(* IEC 61131-3 sources: SemaPLC/sema-plc-benchmark/spec2control-benchmark/data/st-baseline/coking-refinery/pous/programs, 9 files *)

(* ---- main.st ---- *)
PROGRAM main
VAR
	Heartbeat : bool;
END_VAR

(* Entry point required by OpenPLC Editor v4. The process sections run as parallel program instances under task0; main only provides a scan heartbeat. *)
Heartbeat := NOT Heartbeat;

END_PROGRAM

(* ---- Section2.st ---- *)
PROGRAM Section2
VAR
	FT101_FeedFlow_PV_kgphr : real;
	FT102_RefluxFlow_PV_kgphr : real;
	FFIC103_RefluxFlow_SP_kgphr : real;
	FIC104_Output_Percent : real;
	FV104_ValvePosition_Percent : real;
	FV104_FeedbackPos_Percent : real;
	FV104_ValveMoving : bool;
	PIT106_ColumnPressure_bar : real;
	TIT104_Temperature_C : real;
	TIT105_Temperature_C : real;
	TIT107_Temperature_C : real;
	FT_101 : ANALOG_IN;
	FT_102 : ANALOG_IN;
	PIT_106 : ANALOG_IN;
	TIT_104 : ANALOG_IN;
	TIT_105 : ANALOG_IN;
	TIT_107 : ANALOG_IN;
	FFIC_103 : RATIO_CONTROL;
	FIC_104 : PID_BASIC;
	FV_104 : VALVE_ELECTRIC;
	RatioInhibit_OR : bool;
	FeedNotAbove500_NOT : bool;
	ValveInhibit_OR : bool;
END_VAR

FT_101(
    PV_Low := 100.0,
    Scaling_Slope := 312.5,
    Scaling_Offset := -1250.0,
    Alarm_Enable := TRUE);
FT_102(
    Scaling_Slope := 156.25,
    Scaling_Offset := -625.0,
    Alarm_Enable := TRUE);
PIT_106(
    PV_High := 1.5,
    PV_Low := 0.5,
    Alarm_Enable := TRUE);
TIT_104(
    PV_High := 350.0,
    PV_Low := 120.0,
    Alarm_Enable := TRUE);
TIT_105(
    PV_High := 350.0,
    PV_Low := 120.0,
    Alarm_Enable := TRUE);
TIT_107(
    PV_High := 350.0,
    PV_Low := 120.0,
    Alarm_Enable := TRUE);
FIC_104(
    AUTO := TRUE,
    PV := FT_102.PV,
    SP := FFIC_103.SlaveSP,
    MV_MIN := 0.0,
    MV_MAX := 100.0,
    Inhibit := RatioInhibit_OR);
FeedNotAbove500_NOT := NOT FT_101.High_Alarm;
ValveInhibit_OR := FeedNotAbove500_NOT OR TIT_104.High_Alarm OR TIT_104.Low_Alarm OR TIT_105.High_Alarm OR TIT_105.Low_Alarm OR TIT_107.High_Alarm OR TIT_107.Low_Alarm;
FV_104(
    Control_Signal := FIC_104.XOUT,
    Manual_Mode := FALSE,
    Open_Limit := 100.0,
    Close_Limit := 0.0,
    Inhibit := ValveInhibit_OR);
RatioInhibit_OR := PIT_106.High_Alarm OR PIT_106.Low_Alarm OR TIT_104.High_Alarm OR TIT_104.Low_Alarm OR TIT_105.High_Alarm OR TIT_105.Low_Alarm OR TIT_107.High_Alarm OR TIT_107.Low_Alarm OR FT_101.Low_Alarm OR FT_101.General_Fault OR FT_102.General_Fault OR FV_104.Position_Error;
FFIC_103(
    Auto := TRUE,
    PrimaryPV := FT_101.PV,
    SecondaryPV := FT_102.PV,
    RatioSP := 0.5,
    Bias := 0.0,
    MV_MIN := 0.0,
    MV_MAX := 2500.0,
    Inhibit := RatioInhibit_OR);

(* Outputs published to other sections / HMI. *)
FT101_FeedFlow_PV_kgphr := FT_101.PV;
FT102_RefluxFlow_PV_kgphr := FT_102.PV;
FFIC103_RefluxFlow_SP_kgphr := FFIC_103.SlaveSP;
FIC104_Output_Percent := FIC_104.XOUT;
FV104_ValvePosition_Percent := FV_104.Valve_Position;
FV104_FeedbackPos_Percent := FV_104.Feedback_Pos;
FV104_ValveMoving := FV_104.Valve_Moving;
PIT106_ColumnPressure_bar := PIT_106.PV;
TIT104_Temperature_C := TIT_104.PV;
TIT105_Temperature_C := TIT_105.PV;
TIT107_Temperature_C := TIT_107.PV;

END_PROGRAM

(* ---- Section3.st ---- *)
PROGRAM Section3
VAR
	PIT_103_PV_mmHg : real;
	PIC_102_MV_Percent : real;
	PIT_103 : ANALOG_IN;
	PIC_102 : PID_BASIC;
	PV_101 : VALVE_ELECTRIC;
	VDU_START_OK : BOOL_INPUT;
	MAINT_BYPASS_OK : BOOL_INPUT;
	PIC102Inhibit_OR : bool;
	PV101Inhibit_OR : bool;
	VDUStartPermissive_NOT : bool;
END_VAR

PIT_103(
    PV_High := 80.0,
    PV_Low := 20.0,
    Scaling_Slope := 47.5,
    Scaling_Offset := -190.0,
    Alarm_Enable := TRUE);
MAINT_BYPASS_OK();
VDU_START_OK();
VDUStartPermissive_NOT := NOT VDU_START_OK.Bool_Out;
PIC102Inhibit_OR := VDUStartPermissive_NOT OR MAINT_BYPASS_OK.Bool_Out OR PIT_103.General_Fault OR PIC_102.PV_Low_Alarm;
PIC_102(
    AUTO := TRUE,
    PV := PIT_103.PV,
    SP := 50.0,
    MV_MIN := 0.0,
    MV_MAX := 100.0,
    KP := 1.8,
    TR := 2.0,
    TD := 0.5,
    Deviation_Limit := 5.0,
    Inhibit := PIC102Inhibit_OR);
PV101Inhibit_OR := PIC_102.PV_High_Alarm OR PV_101.Position_Error;
PV_101(
    Control_Signal := PIC_102.XOUT,
    Open_Limit := 100.0,
    Close_Limit := 0.0,
    Inhibit := PV101Inhibit_OR);

(* Outputs published to other sections / HMI. *)
PIT_103_PV_mmHg := PIT_103.PV;
PIC_102_MV_Percent := PIC_102.XOUT;

END_PROGRAM

(* ---- Section4.st ---- *)
PROGRAM Section4
VAR
	PC301_SP_Operator : real;
	PT_301_RegeneratorPressure_PV : real;
	PT_302_BlowerDischargePressure_PV : real;
	PT_303_FractionatorOverheadPressure_PV : real;
	TT_301_RegeneratorTemperature_PV : real;
	PTF_301_FilteredPressure_PV : real;
	PC_301_Output_to_PV_105_Percent : real;
	PV_105_Valve_Position_Command_Percent : real;
	PV_105_Valve_Position_Feedback_Percent : real;
	P_301A_Running_Status : bool;
	XV_108_Closed_Status : bool;
	PT_301 : ANALOG_IN;
	PT_302 : ANALOG_IN;
	PT_303 : ANALOG_IN;
	PTF_301 : ANALOG_IN;
	TT_301 : ANALOG_IN;
	PC_301 : PID_BASIC;
	PV_105 : VALVE_ELECTRIC;
	PV_106 : VALVE_ON_OFF;
	XV_108 : VALVE_ON_OFF;
	P_301A : MOTOR_ON_OFF;
	SteadyState_TON : TON;
	SetpointClamp_LIMIT : real;
	StartupSP_Select_SEL : real;
	ErrorCalc_SUB : real;
	ErrorPos_GT : bool;
	ErrorNeg_LT : bool;
	ErrorOutsideBand_OR : bool;
	DeadbandApply_SEL : real;
	PV_Reconstruct_ADD : real;
	BlowerNotRunning_NOT : bool;
	Permissives_OR1 : bool;
	Permissives_OR2 : bool;
	Permissives_OR3 : bool;
	PV105Inhibit_OR : bool;
	AutoHold_OR : bool;
	AutoEnable_NOT : bool;
	ESD_HighPressure_GT : bool;
	ReliefValve_GT : bool;
	ReliefValve_Close_NOT : bool;
	OutsideBand_NOT : bool;
END_VAR

PT_301(
    PV_High := 2.8,
    PV_Low := 2.2,
    Scaling_Slope := 0.3125,
    Scaling_Offset := -1.25,
    Alarm_Enable := TRUE);
PT_302(
    Scaling_Slope := 0.3125,
    Scaling_Offset := -1.25,
    Alarm_Enable := TRUE);
PT_303(
    Scaling_Slope := 0.3125,
    Scaling_Offset := -1.25,
    Alarm_Enable := TRUE);
PTF_301(
    Scaling_Slope := 0.3125,
    Scaling_Offset := -1.25);
TT_301(
    Scaling_Slope := 62.5,
    Scaling_Offset := -250.0,
    Alarm_Enable := TRUE);
ESD_HighPressure_GT := (PT_301.PV > 3.0);
XV_108(
    Open_Cmd := FALSE,
    Close_Cmd := ESD_HighPressure_GT,
    Timeout := T#5s);
AutoHold_OR := PT_301.General_Fault OR XV_108.FB_Closed;
AutoEnable_NOT := NOT AutoHold_OR;
ErrorNeg_LT := (ErrorCalc_SUB < -0.05);
ErrorPos_GT := (ErrorCalc_SUB > 0.05);
ErrorOutsideBand_OR := ErrorPos_GT OR ErrorNeg_LT;
OutsideBand_NOT := NOT ErrorOutsideBand_OR;
SteadyState_TON(
    IN := OutsideBand_NOT,
    PT := T#60s);
StartupSP_Select_SEL := SEL(G := SteadyState_TON.Q, IN0 := 2.5, IN1 := 0.0);
ErrorCalc_SUB := PT_301.PV - StartupSP_Select_SEL;
DeadbandApply_SEL := SEL(G := ErrorOutsideBand_OR, IN0 := 0.0, IN1 := ErrorCalc_SUB);
PV_Reconstruct_ADD := StartupSP_Select_SEL + DeadbandApply_SEL;
PC_301(
    AUTO := AutoEnable_NOT,
    PV := PV_Reconstruct_ADD,
    SP := StartupSP_Select_SEL,
    MV_MIN := 0.0,
    MV_MAX := 100.0,
    X0 := 0.0,
    KP := 3.0,
    TR := 1.2,
    TD := 0.1);
P_301A();
BlowerNotRunning_NOT := NOT P_301A.FB_Running;
Permissives_OR1 := TT_301.Low_Alarm OR BlowerNotRunning_NOT;
Permissives_OR2 := PT_302.Low_Alarm OR PT_303.High_Alarm;
Permissives_OR3 := Permissives_OR1 OR Permissives_OR2;
PV105Inhibit_OR := Permissives_OR3 OR XV_108.FB_Closed;
PV_105(
    Control_Signal := PC_301.XOUT,
    Manual_Mode := FALSE,
    Open_Limit := 100.0,
    Close_Limit := 0.0,
    Timeout := T#10s,
    Inhibit := PV105Inhibit_OR);
ReliefValve_GT := (PT_301.PV > 3.5);
ReliefValve_Close_NOT := NOT ReliefValve_GT;
PV_106(
    Open_Cmd := ReliefValve_GT,
    Close_Cmd := ReliefValve_Close_NOT,
    Timeout := T#5s);
SetpointClamp_LIMIT := LIMIT(MN := 2.0, IN := PC301_SP_Operator, MX := 3.0);

(* Outputs published to other sections / HMI. *)
PT_301_RegeneratorPressure_PV := PT_301.PV;
PT_302_BlowerDischargePressure_PV := PT_302.PV;
PT_303_FractionatorOverheadPressure_PV := PT_303.PV;
TT_301_RegeneratorTemperature_PV := TT_301.PV;
PTF_301_FilteredPressure_PV := PTF_301.PV;
PC_301_Output_to_PV_105_Percent := PC_301.XOUT;
PV_105_Valve_Position_Command_Percent := PV_105.Valve_Position;
PV_105_Valve_Position_Feedback_Percent := PV_105.Feedback_Pos;
P_301A_Running_Status := P_301A.FB_Running;
XV_108_Closed_Status := XV_108.FB_Closed;

END_PROGRAM

(* ---- Section5.st ---- *)
PROGRAM Section5
VAR
	TIT101_FurnaceOutletTemp_PV_C : real;
	TC401_FV401_FuelGas_MV_Pct : real;
	PT402_FurnaceDraft_PV_kPa : real;
	PT403_DischargePressure_PV_bar : real;
	PC401_FuelGasPressure_PV_bar : real;
	TIT101_HighTempAlarm_3s : bool;
	TIT101_LowTempAlarm_3s : bool;
	TIT_101 : ANALOG_IN;
	TC_401 : PID_BASIC;
	FV_401 : VALVE_ELECTRIC;
	PT_402 : ANALOG_IN;
	PT_403 : ANALOG_IN;
	PC_401 : PID_BASIC;
	FT_401A : DIGITAL_IN;
	FT_401B : DIGITAL_IN;
	FuelGasInterlockDelay_TON : TON;
	TIT101_HighAlarmDelay_TON : TON;
	TIT101_LowAlarmDelay_TON : TON;
	FlameLitPermissive_AND : bool;
	FlameNotLit_NOT : bool;
	FuelGasPermissiveViolations_OR : bool;
	MasterInhibit_OR : bool;
END_VAR

TIT_101(
    PV_High := 510.0,
    PV_Low := 480.0,
    Scaling_Slope := 9.375,
    Scaling_Offset := 362.5,
    Alarm_Enable := TRUE);
FT_401A();
FT_401B();
FlameLitPermissive_AND := FT_401A.DI_Out AND FT_401B.DI_Out;
FlameNotLit_NOT := NOT FlameLitPermissive_AND;
PC_401(
    PV := PC401_FuelGasPressure_PV_bar);
PT_402(
    Alarm_Enable := TRUE);
PT_403(
    Alarm_Enable := TRUE);
FuelGasPermissiveViolations_OR := PC_401.PV_High_Alarm OR PC_401.PV_Low_Alarm OR PT_402.High_Alarm OR PT_402.Low_Alarm OR PT_403.Low_Alarm;
FuelGasInterlockDelay_TON(
    IN := FuelGasPermissiveViolations_OR,
    PT := T#5s);
MasterInhibit_OR := TC_401.PV_High_Alarm OR FuelGasInterlockDelay_TON.Q OR FlameNotLit_NOT OR TIT_101.General_Fault;
FV_401(
    Control_Signal := TC_401.XOUT,
    Manual_Mode := FALSE,
    Open_Limit := 100.0,
    Close_Limit := 0.0,
    Inhibit := MasterInhibit_OR);
TC_401(
    AUTO := TRUE,
    PV := TIT_101.PV,
    SP := 495.0,
    MV_MIN := 0.0,
    MV_MAX := 100.0,
    X0 := FV_401.Feedback_Pos,
    KP := 3.2,
    TR := 0.9,
    TD := 0.3,
    Deviation_Limit := 2.0,
    Inhibit := MasterInhibit_OR);
TIT101_HighAlarmDelay_TON(
    IN := TIT_101.High_Alarm,
    PT := T#3s);
TIT101_LowAlarmDelay_TON(
    IN := TIT_101.Low_Alarm,
    PT := T#3s);

(* Outputs published to other sections / HMI. *)
TIT101_FurnaceOutletTemp_PV_C := TIT_101.PV;
TC401_FV401_FuelGas_MV_Pct := TC_401.XOUT;
PT402_FurnaceDraft_PV_kPa := PT_402.PV;
PT403_DischargePressure_PV_bar := PT_403.PV;
TIT101_HighTempAlarm_3s := TIT101_HighAlarmDelay_TON.Q;
TIT101_LowTempAlarm_3s := TIT101_LowAlarmDelay_TON.Q;

END_PROGRAM

(* ---- Section6.st ---- *)
PROGRAM Section6
VAR
	FT103_H2Flow_PV : real;
	FC103_MV_Percent : real;
	TT101_Temp_PV : real;
	TC501_MV_Percent : real;
	PT501_Pressure_PV : real;
	PT502_InletPressure_PV : real;
	FC103_SP_Operator : real;
	FC103_SP_Clamped : real;
	FC103_SP_Reduced : real;
	FT_103 : ANALOG_IN;
	FC_103 : PID_BASIC;
	FV_103 : VALVE_ELECTRIC;
	TT_101 : ANALOG_IN;
	TC_501 : PID_BASIC;
	TV_501 : VALVE_ELECTRIC;
	PT_501 : ANALOG_IN;
	PC_501 : PID_BASIC;
	PT_502 : ANALOG_IN;
	ESD_501 : DIGITAL_IN;
	TV501_OpenDelay_TON : TON;
	FC103_Inhibit_OR : bool;
	TV501_Inhibit_OR : bool;
	TC501_Inhibit_OR : bool;
	PT501_OverLimit_GT : bool;
	FC103_SP_Half_MULT : real;
	FC103_SP_SEL : real;
	H2_Shutdown_OR : bool;
	H2_Auto_NOT : bool;
	ESD_NOT : bool;
	PT502_Permissive_GT : bool;
	TV501_Permissive_AND : bool;
	TV501_AutoReady_NOT : bool;
	TV501_ManualMode_OR : bool;
	TV501_ManualPos_SEL : real;
	FC103_SP_Max_MAX : real;
	FC103_SP_Clamp_MIN : real;
END_VAR

FT_103(
    Scaling_Slope := 125.0,
    Scaling_Offset := -500.0,
    Alarm_Enable := TRUE);
ESD_501();
TT_101(
    Alarm_Enable := TRUE);
FC103_Inhibit_OR := ESD_501.DI_Out OR TT_101.High_Alarm OR FT_103.General_Fault;
FC103_SP_Max_MAX := MAX(FC103_SP_Operator, 500.0);
FC103_SP_Clamp_MIN := MIN(FC103_SP_Max_MAX, 1500.0);
FC103_SP_Half_MULT := FC103_SP_Clamp_MIN * 0.5;
PT_501();
PT501_OverLimit_GT := (PT_501.PV > 50.0);
FC103_SP_SEL := SEL(G := PT501_OverLimit_GT, IN0 := FC103_SP_Clamp_MIN, IN1 := FC103_SP_Half_MULT);
H2_Shutdown_OR := ESD_501.DI_Out OR TT_101.High_Alarm;
H2_Auto_NOT := NOT H2_Shutdown_OR;
FC_103(
    AUTO := H2_Auto_NOT,
    PV := FT_103.PV,
    SP := FC103_SP_SEL,
    MV_MIN := 0.0,
    MV_MAX := 100.0,
    KP := 1.8,
    TR := 0.5,
    TD := 0.1,
    PV_High := 1600.0,
    PV_Low := 400.0,
    Inhibit := FC103_Inhibit_OR);
FV_103(
    Control_Signal := FC_103.XOUT,
    Manual_Mode := H2_Shutdown_OR,
    Open_Limit := 100.0,
    Close_Limit := 0.0,
    Inhibit := FC103_Inhibit_OR);
ESD_NOT := NOT ESD_501.DI_Out;
TC501_Inhibit_OR := ESD_501.DI_Out OR TT_101.General_Fault;
TC_501(
    AUTO := ESD_NOT,
    PV := TT_101.PV,
    SP := 375.0,
    MV_MIN := 0.0,
    MV_MAX := 100.0,
    KP := 2.5,
    TR := 0.8,
    TD := 0.2,
    PV_High := 415.0,
    PV_Low := 290.0,
    Inhibit := TC501_Inhibit_OR);
PT_502(
    Alarm_Enable := TRUE);
TV501_Inhibit_OR := ESD_501.DI_Out OR PT_502.Low_Alarm OR TT_101.General_Fault;
PT502_Permissive_GT := (PT_502.PV > 10.0);
TV501_Permissive_AND := ESD_NOT AND PT502_Permissive_GT;
TV501_OpenDelay_TON(
    IN := TV501_Permissive_AND,
    PT := T#15s);
TV501_AutoReady_NOT := NOT TV501_OpenDelay_TON.Q;
TV501_ManualMode_OR := TV501_AutoReady_NOT OR ESD_501.DI_Out;
TV501_ManualPos_SEL := SEL(G := ESD_501.DI_Out, IN0 := 0.0, IN1 := 100.0);
TV_501(
    Control_Signal := TC_501.XOUT,
    Manual_Mode := TV501_ManualMode_OR,
    Manual_Position := TV501_ManualPos_SEL,
    Open_Limit := 100.0,
    Close_Limit := 0.0,
    Inhibit := TV501_Inhibit_OR);
PC_501(
    PV := PT_501.PV,
    Inhibit := ESD_501.DI_Out);

(* Outputs published to other sections / HMI. *)
FT103_H2Flow_PV := FT_103.PV;
FC103_MV_Percent := FC_103.XOUT;
TT101_Temp_PV := TT_101.PV;
TC501_MV_Percent := TC_501.XOUT;
PT501_Pressure_PV := PT_501.PV;
PT502_InletPressure_PV := PT_502.PV;

END_PROGRAM

(* ---- Section7.st ---- *)
PROGRAM Section7
VAR
	FT601_Raw_mA : real;
	LT601_Raw_mA : real;
	TT104_Raw_mA : real;
	FT601_FlowRate_m3h_PV : real;
	LT601_SiloLevel_Pct_PV : real;
	TT104_Temperature_C_PV : real;
	FIC601_MV_Pct : real;
	P601A_SpeedCmd_Pct : real;
	P601B_SpeedCmd_Pct : real;
	SP_Operator_m3h : real;
	FA601_LowFlow_Alarm : bool;
	LAH601_HighLevel_Alarm : bool;
	TAH104_HighTemp_Alarm : bool;
	Start_Pumps_Cmd : bool;
	Stop_Pumps_Cmd : bool;
	MCC601_Status_In : bool;
	MCC602_Status_In : bool;
	Crusher_RunPermissive : bool;
	Permissive_All_OK : bool;
	FT601_Signal_OK : bool;
	FT_601 : ANALOG_IN;
	LT_601 : ANALOG_IN;
	TT_104 : ANALOG_IN;
	FIC_601 : PID_BASIC;
	P_601A : MOTOR_VSD;
	P_601B : MOTOR_VSD;
	MCC_601 : BOOL_INPUT;
	MCC_602 : BOOL_INPUT;
	StartDelay_TON : TON;
	LowFlowDelay_TON : TON;
	PumpsInhibit_OR : bool;
	LevelPermissive_GE : bool;
	TempPermissive_LE : bool;
	PumpsPermissive_AND : bool;
	FT601Fault_NOT : bool;
	LowFlow_LT : bool;
	PumpA_Start_AND : bool;
	PumpB_Start_AND : bool;
	PumpA_Stop_OR : bool;
	B_StartSource_OR : bool;
	CrusherPermissive_AND : bool;
	SP_ClampHigh_MIN : real;
	SP_ClampLow_MAX : real;
	HighLevel_LT601_GT : bool;
END_VAR

FT_601(
    Raw_Signal := FT601_Raw_mA,
    PV_Low := 80.0,
    Scaling_Slope := 15.625,
    Scaling_Offset := -62.5,
    Alarm_Enable := TRUE);
LT_601(
    Raw_Signal := LT601_Raw_mA,
    PV_High := 90.0,
    Scaling_Slope := 6.25,
    Scaling_Offset := -25.0,
    Alarm_Enable := TRUE);
TT_104(
    Raw_Signal := TT104_Raw_mA,
    PV_High := 85.0,
    Scaling_Slope := 6.25,
    Scaling_Offset := -25.0,
    Alarm_Enable := TRUE);
FT601Fault_NOT := NOT FT_601.General_Fault;
SP_ClampHigh_MIN := MIN(SP_Operator_m3h, 200.0);
SP_ClampLow_MAX := MAX(SP_ClampHigh_MIN, 100.0);
FIC_601(
    AUTO := FT601Fault_NOT,
    PV := FT_601.PV,
    SP := SP_ClampLow_MAX,
    MV_MIN := 20.0,
    MV_MAX := 100.0,
    X0 := 0.0,
    KP := 2.0,
    TR := 1.5,
    TD := 0.3,
    Inhibit := FT_601.General_Fault);
LevelPermissive_GE := (LT_601.PV >= 10.0);
TempPermissive_LE := (TT_104.PV <= 80.0);
PumpsPermissive_AND := LevelPermissive_GE AND TempPermissive_LE;
StartDelay_TON(
    IN := PumpsPermissive_AND,
    PT := T#5s);
PumpA_Start_AND := Start_Pumps_Cmd AND StartDelay_TON.Q;
PumpsInhibit_OR := LT_601.Low_Alarm OR TT_104.High_Alarm;
PumpA_Stop_OR := PumpsInhibit_OR OR Stop_Pumps_Cmd;
P_601A(
    Start_Cmd := PumpA_Start_AND,
    Stop_Cmd := PumpA_Stop_OR,
    Speed_SP := FIC_601.XOUT,
    Accel_Ramp := T#2s,
    Decel_Ramp := T#2s,
    Inhibit := PumpsInhibit_OR);
B_StartSource_OR := P_601A.FB_Fault OR Start_Pumps_Cmd;
PumpB_Start_AND := B_StartSource_OR AND StartDelay_TON.Q;
P_601B(
    Start_Cmd := PumpB_Start_AND,
    Stop_Cmd := PumpA_Stop_OR,
    Speed_SP := FIC_601.XOUT,
    Accel_Ramp := T#2s,
    Decel_Ramp := T#2s,
    Inhibit := PumpsInhibit_OR);
MCC_601(
    Bool_In := MCC601_Status_In);
MCC_602(
    Bool_In := MCC602_Status_In);
LowFlow_LT := (FT_601.PV < 80.0);
LowFlowDelay_TON(
    IN := LowFlow_LT,
    PT := T#10s);
CrusherPermissive_AND := MCC_601.Bool_Out AND MCC_602.Bool_Out;
HighLevel_LT601_GT := (LT_601.PV > 90.0);

(* Outputs published to other sections / HMI. *)
FT601_FlowRate_m3h_PV := FT_601.PV;
LT601_SiloLevel_Pct_PV := LT_601.PV;
TT104_Temperature_C_PV := TT_104.PV;
FIC601_MV_Pct := FIC_601.XOUT;
Permissive_All_OK := StartDelay_TON.Q;
Crusher_RunPermissive := CrusherPermissive_AND;
P601A_SpeedCmd_Pct := P_601A.Speed_Out;
P601B_SpeedCmd_Pct := P_601B.Speed_Out;
FA601_LowFlow_Alarm := LowFlowDelay_TON.Q;
LAH601_HighLevel_Alarm := HighLevel_LT601_GT;
TAH104_HighTemp_Alarm := TT_104.High_Alarm;
FT601_Signal_OK := FT601Fault_NOT;

END_PROGRAM

(* ---- Section8.st ---- *)
PROGRAM Section8
VAR
	FT702_AirFlow_SP : real;
	FT_701 : ANALOG_IN;
	FT_702 : ANALOG_IN;
	PT_701 : ANALOG_IN;
	FD_701 : BOOL_INPUT;
	FFIC_701 : RATIO_CONTROL;
	FIC_702 : PID_BASIC;
	LIC_101 : PID_BASIC;
	FV_701 : VALVE_ELECTRIC;
	FV_702 : VALVE_ELECTRIC;
	FlameNotProven_NOT : bool;
	FFIC701_Inhibit_OR : bool;
	FIC702_Inhibit_OR : bool;
	FV701_Inhibit_OR : bool;
	FV702_Inhibit_OR : bool;
END_VAR

FT_701(
    PV_High := 450.0,
    PV_Low := 50.0,
    Alarm_Enable := TRUE);
FT_702(
    Alarm_Enable := TRUE);
PT_701(
    Alarm_Enable := TRUE);
FD_701();
LIC_101();
FV701_Inhibit_OR := LIC_101.PV_High_Alarm OR LIC_101.PV_Low_Alarm OR PT_701.Low_Alarm;
FlameNotProven_NOT := NOT FD_701.Bool_Out;
FFIC701_Inhibit_OR := FlameNotProven_NOT OR FV701_Inhibit_OR OR FT_701.General_Fault OR FT_702.General_Fault;
FFIC_701(
    Auto := TRUE,
    PrimaryPV := FT_701.PV,
    SecondaryPV := FT_702.PV,
    RatioSP := 10.0,
    Bias := 0.0,
    MV_MIN := 500.0,
    MV_MAX := 5000.0,
    ManOut := 2500.0,
    Inhibit := FFIC701_Inhibit_OR);
FIC702_Inhibit_OR := FV701_Inhibit_OR OR FT_701.General_Fault OR FT_702.General_Fault;
FIC_702(
    AUTO := TRUE,
    PV := FT_702.PV,
    SP := FFIC_701.SlaveSP,
    MV_MIN := 0.0,
    MV_MAX := 100.0,
    Deviation_Limit := 500.0,
    Inhibit := FIC702_Inhibit_OR);
FV_701(
    Inhibit := FV701_Inhibit_OR);
FV702_Inhibit_OR := FV701_Inhibit_OR OR FT_701.Low_Alarm;
FV_702(
    Control_Signal := FIC_702.XOUT,
    Inhibit := FV702_Inhibit_OR);

(* Outputs published to other sections / HMI. *)
FT702_AirFlow_SP := FFIC_701.SlaveSP;

END_PROGRAM

(* ---- Section9.st ---- *)
PROGRAM Section9
VAR
	PT106_PV_Pct : real;
	PIC101_MV_Pct : real;
	FV102_Feedback_Pos_Pct : real;
	PT_106 : ANALOG_IN;
	PIC_101 : PID_BASIC;
	FV_102 : VALVE_ELECTRIC;
	LC_801_LEVEL_OK : BOOL_INPUT;
	FLARE_IGNITION_OK : BOOL_INPUT;
	PT_106_VALID : BOOL_INPUT;
	FlareIgnitionFail_NOT : bool;
	PT106_Invalid_NOT : bool;
	PIC101_Inhibit_OR : bool;
	LevelNotOK_NOT : bool;
	FV102_Inhibit_OR : bool;
	DeadbandHold_SEL : real;
END_VAR

PT_106(
    Scaling_Slope := 0.3125,
    Scaling_Offset := -1.25,
    Alarm_Enable := TRUE);
DeadbandHold_SEL := SEL(G := PIC_101.Deviation_Alarm, IN0 := FV_102.Feedback_Pos, IN1 := PIC_101.XOUT);
LC_801_LEVEL_OK();
LevelNotOK_NOT := NOT LC_801_LEVEL_OK.Bool_Out;
FV102_Inhibit_OR := LevelNotOK_NOT OR PIC_101.PV_High_Alarm OR PIC_101.PV_Low_Alarm;
FV_102(
    Control_Signal := DeadbandHold_SEL,
    Open_Limit := 100.0,
    Close_Limit := 0.0,
    Inhibit := FV102_Inhibit_OR);
FLARE_IGNITION_OK();
FlareIgnitionFail_NOT := NOT FLARE_IGNITION_OK.Bool_Out;
PT_106_VALID();
PT106_Invalid_NOT := NOT PT_106_VALID.Bool_Out;
PIC101_Inhibit_OR := FlareIgnitionFail_NOT OR FV_102.Position_Error OR PT106_Invalid_NOT OR PT_106.General_Fault;
PIC_101(
    AUTO := TRUE,
    PV := PT_106.PV,
    SP := 1.5,
    MV_MIN := 0.0,
    MV_MAX := 100.0,
    X0 := FV_102.Feedback_Pos,
    KP := -3.2,
    TR := 0.5,
    TD := 0.1,
    PV_High := 1.8,
    PV_Low := 1.2,
    Deviation_Limit := 0.15,
    Inhibit := PIC101_Inhibit_OR);

(* Outputs published to other sections / HMI. *)
PT106_PV_Pct := PT_106.PV;
PIC101_MV_Pct := PIC_101.XOUT;
FV102_Feedback_Pos_Pct := FV_102.Feedback_Pos;

END_PROGRAM
